Fanuc KAREL source: KA00109.KL

PROGRAM KA00109
%NOLOCKGROUP
VAR
  SRC: CONFIG
  DST: INTEGER
BEGIN
  SRC.CFG_FLIP = TRUE
  DST = SRC
END KA00109
